//{attribute 'qualified_only'}
VAR_GLOBAL
    {attribute 'pytmc' :=' pv: RTDSL0:MPA:01 '}
    RTDSL0_MPA_01: FB_MPA := (sName := 'RTDSL0:MPA:01');

    {attribute 'pytmc' :=' pv: RTDSL0:MPA:02 '}
    RTDSL0_MPA_02: FB_MPA := (sName := 'RTDSL0:MPA:02');

    {attribute 'pytmc' :=' pv: RTDSL0:MPA:03 '}
    RTDSL0_MPA_03: FB_MPA := (sName := 'RTDSL0:MPA:03');

    {attribute 'pytmc' :=' pv: RTDSL0:MPA:04 '}
    RTDSL0_MPA_04: FB_MPA := (sName := 'RTDSL0:MPA:04');


END_VAR

(* stored: Version 1.1.0.1, ProductVersion 3.1.4022.18
   GVL RTDSL0: Id {ac721235-6abd-4ba5-afeb-f19d34581d05} *)
